Staubli VAL3: copyItem.pgx

public program copyItem(string x_sTarget, string x_sSource)
  local num l_nSize
  local num l_i
  local num l_j
begin
  l_nSize=size(progTemp:pProgItem[x_sSource].pProgTemplate)
  resize(progTemp:pProgItem[x_sTarget].pProgTemplate,1,l_nSize)
  for l_i = 0 to l_nSize-1
    progTemp:pProgItem[x_sTarget].pProgTemplate[l_i].sTRAJname=progTemp:pProgItem[x_sSource].pProgTemplate[l_i].sTRAJname
    progTemp:pProgItem[x_sTarget].pProgTemplate[l_i].nType=progTemp:pProgItem[x_sSource].pProgTemplate[l_i].nType
    for l_j=0 to 2
      progTemp:pProgItem[x_sTarget].pProgTemplate[l_i].iIfItem.nSigType[l_j]=progTemp:pProgItem[x_sSource].pProgTemplate[l_i].iIfItem.nSigType[l_j]
      progTemp:pProgItem[x_sTarget].pProgTemplate[l_i].iIfItem.nSigIndex[l_j]=progTemp:pProgItem[x_sSource].pProgTemplate[l_i].iIfItem.nSigIndex[l_j]
      progTemp:pProgItem[x_sTarget].pProgTemplate[l_i].iIfItem.nValue[l_j]=progTemp:pProgItem[x_sSource].pProgTemplate[l_i].iIfItem.nValue[l_j]
    endFor
    progTemp:pProgItem[x_sTarget].pProgTemplate[l_i].iIfItem.bANDOR[0]=(progTemp:pProgItem[x_sSource].pProgTemplate[l_i].iIfItem.bANDOR[0]==true)
    progTemp:pProgItem[x_sTarget].pProgTemplate[l_i].iIfItem.bANDOR[1]=(progTemp:pProgItem[x_sSource].pProgTemplate[l_i].iIfItem.bANDOR[1]==true)
  endFor
end
